TYPE "ST_DeclarationParCfg"
VERSION : 0.1
   STRUCT
      SchemaVersion : UInt := 4;
      Timeout : Time := T#8S;
      Preset : DInt := 10;
   END_STRUCT;

END_TYPE

